Staubli VAL3: safeData.pjx

--- safeData.pjx ---
Parameters version=s8.10.3Cs9_BS2093 stackSize=5000 millimeterUnit=true
Program file=start.pgx
Program file=stop.pgx
Data file=safeData.dtx
Type name=zoneItem path=Disk://source/template/zoneTemplate/zoneTemplate.pjx
Type name=sPoint path=Disk://source/template/sPointTemplate/sPointTemplate.pjx

--- safeData.dtx ---
public sPoint sSPoint[16]
  [0]
    bool bActive = true
    pointRx pPointRx = {x=749.14032, y=226.565031, z=1244.301358, rx=-64.150648, ry=3.461024, rz=92.316205, shoulder=lefty, elbow=enegative, wrist=wpositive, fatherId=world[0]}
    string sName = "安全点0"
  [1]
    bool bActive = true
    pointRx pPointRx = {x=749.140309, y=226.565029, z=1244.301359, rx=-64.150648, ry=3.461022, rz=92.316204, shoulder=lefty, elbow=enegative, wrist=wpositive, fatherId=world[0]}
    string sName = "安全点1"
  [2]
    bool bActive
    pointRx pPointRx
    string sName = "安全点2"
  [3]
    bool bActive
    pointRx pPointRx
    string sName = "安全点3"
  [4]
    bool bActive = true
    pointRx pPointRx = {x=1166.518639, y=208.558661, z=446.0719177, rx=49.817861, ry=102.228281, rz=-47.114554, shoulder=lefty, elbow=epositive, wrist=wnegative, fatherId=world[0]}
    string sName = "安全点4"
  [5]
    bool bActive = true
    pointRx pPointRx = {x=1166.518639, y=208.558696, z=446.0719088, rx=49.81785, ry=102.228285, rz=-47.11454, shoulder=lefty, elbow=epositive, wrist=wnegative, fatherId=world[0]}
    string sName = "安全点5"
  [6]
    bool bActive
    pointRx pPointRx
    string sName = "安全点6"
  [7]
    bool bActive
    pointRx pPointRx
    string sName = "安全点7"
  [8]
    bool bActive
    pointRx pPointRx
    string sName = "安全点8"
  [9]
    bool bActive
    pointRx pPointRx
    string sName = "安全点9"
  [10]
    bool bActive
    pointRx pPointRx
    string sName
  [11]
    bool bActive
    pointRx pPointRx
    string sName
  [12]
    bool bActive
    pointRx pPointRx
    string sName
  [13]
    bool bActive
    pointRx pPointRx
    string sName
  [14]
    bool bActive
    pointRx pPointRx
    string sName
  [15]
    bool bActive
    pointRx pPointRx
    string sName
public zoneItem zZoneItem[16]
  [0]
    bool bActive
    frame fBase = {}
    pointRx pFirst = {shoulder=lefty, elbow=epositive, wrist=wpositive}
    pointRx pO
    pointRx pSecond
    pointRx pX
    pointRx pY
    string sID = "rrff"
  [1]
    bool bActive = true
    frame fBase = {}
    pointRx pFirst = {x=-118.432053, y=-40.166607, z=722.0958456, rx=-35.377493, ry=-42.132282, rz=-101, shoulder=righty, elbow=epositive, wrist=wnegative}
    pointRx pO
    pointRx pSecond = {x=500, y=-1000, z=1000, rx=-35, ry=-42, rz=-100}
    pointRx pX
    pointRx pY
    string sID = "干涉区1"
  [2]
    bool bActive
    frame fBase = {}
    pointRx pFirst
    pointRx pO
    pointRx pSecond
    pointRx pX
    pointRx pY
    string sID = "干涉区2"
  [3]
    bool bActive
    frame fBase = {}
    pointRx pFirst
    pointRx pO
    pointRx pSecond
    pointRx pX
    pointRx pY
    string sID = "干涉区3"
  [4]
    bool bActive
    frame fBase = {}
    pointRx pFirst
    pointRx pO
    pointRx pSecond
    pointRx pX
    pointRx pY
    string sID = "干涉区4"
  [5]
    bool bActive
    frame fBase = {}
    pointRx pFirst
    pointRx pO
    pointRx pSecond
    pointRx pX
    pointRx pY
    string sID = "干涉区5"
  [6]
    bool bActive
    frame fBase = {}
    pointRx pFirst
    pointRx pO
    pointRx pSecond
    pointRx pX
    pointRx pY
    string sID = "干涉区6"
  [7]
    bool bActive
    frame fBase = {}
    pointRx pFirst
    pointRx pO
    pointRx pSecond
    pointRx pX
    pointRx pY
    string sID = "干涉区7"
  [8]
    bool bActive
    frame fBase = {}
    pointRx pFirst
    pointRx pO
    pointRx pSecond
    pointRx pX
    pointRx pY
    string sID = "干涉区8"
  [9]
    bool bActive
    frame fBase = {}
    pointRx pFirst
    pointRx pO
    pointRx pSecond
    pointRx pX
    pointRx pY
    string sID = "干涉区9"
  [10]
    bool bActive
    frame fBase = {}
    pointRx pFirst
    pointRx pO
    pointRx pSecond
    pointRx pX
    pointRx pY
    string sID
  [11]
    bool bActive
    frame fBase = {}
    pointRx pFirst
    pointRx pO
    pointRx pSecond
    pointRx pX
    pointRx pY
    string sID
  [12]
    bool bActive
    frame fBase = {}
    pointRx pFirst
    pointRx pO
    pointRx pSecond
    pointRx pX
    pointRx pY
    string sID
  [13]
    bool bActive
    frame fBase = {}
    pointRx pFirst
    pointRx pO
    pointRx pSecond
    pointRx pX
    pointRx pY
    string sID
  [14]
    bool bActive
    frame fBase = {}
    pointRx pFirst
    pointRx pO
    pointRx pSecond
    pointRx pX
    pointRx pY
    string sID
  [15]
    bool bActive
    frame fBase = {}
    pointRx pFirst
    pointRx pO
    pointRx pSecond
    pointRx pX
    pointRx pY
    string sID

--- start.pgx ---
program start()
begin
end

--- stop.pgx ---
program stop()
begin
end
